// TIA Portal V20 export
Screen "190FX1Layout_Docking"  1276x673
  ScreenItem "Line_Header_X0_Y64" at 0,64 size 1276x0  Type=HmiLine
  ScreenItem "permanentareaborderrectangle" at 0,0 size 0x0  Type=HmiRectangle
  ScreenItem "Button_Back" at 2,2 size 90x60  Type=HmiButton
  ScreenItem "Move_Legend" at 1183,2 size 90x60  Type=HmiButton
  ScreenItem "Fusszeile_Button_ManualOPMode1_2" at 188,2 size 90x60  Type=HmiButton
  ScreenItem "文本域_22" at 1130,495 size 104x23  Type=HmiTextBox
  ScreenItem "面板容器_23" at 1177,528 size 96x32  Type=HmiFaceplateContainer
  ScreenItem "面板容器_22" at 1067,528 size 96x32  Type=HmiFaceplateContainer
  ScreenItem "面板容器_2" at 1091,4 size 88x58  Type=HmiFaceplateContainer
  ScreenItem "OPMode1_Blocked" at 1165,6 size 14x14  Type=HmiGraphicView
  ScreenItem "OPMode4_Foreground_Blocked" at 1091,4 size 88x58  Type=HmiGraphicView
  ScreenItem "Fusszeile_Button_ManualOPMode1_1" at 95,2 size 90x60  Type=HmiButton
  ScreenItem "LSicar_Valve8Pos_LeftHomeRightWork_WithPB_3" at 1099,110 size 160x53  Type=HmiFaceplateContainer
  ScreenItem "文本域_5" at 1107,83 size 139x22  Type=HmiTextBox
  ScreenItem "面板容器_15" at 54,347 size 65x43  Type=HmiFaceplateContainer
  ScreenItem "Graphic view_1" at 114,71 size 766x527  Type=HmiGraphicView
  ScreenItem "Line_4" at 527,411 size 146x156  Type=HmiLine
  ScreenItem "Line_5" at 509,439 size 5x185  Type=HmiLine
  ScreenItem "Line_6" at 104,365 size 253x0  Type=HmiLine
  ScreenItem "Line_7" at 406,338 size 1x280  Type=HmiLine
  ScreenItem "面板容器_13" at 613,609 size 142x51  Type=HmiFaceplateContainer
  ScreenItem "面板容器_12" at 312,609 size 142x51  Type=HmiFaceplateContainer
  ScreenItem "Faceplate container_5" at 483,609 size 65x43  Type=HmiFaceplateContainer
  ScreenItem "文本域_19" at 34,328 size 100x20  Type=HmiTextBox
  ScreenItem "文本域_6" at 312,567 size 140x40  Type=HmiTextBox
  ScreenItem "文本域_8" at 1172,-248 size 100x20  Type=HmiTextBox
  ScreenItem "文本域_9" at 1741,-563 size 100x20  Type=HmiTextBox
  ScreenItem "文本域_10" at 2310,-878 size 100x20  Type=HmiTextBox
  ScreenItem "文本域_11" at 462,587 size 100x20  Type=HmiTextBox
  ScreenItem "文本域_12" at 321,1215 size 100x20  Type=HmiTextBox
  ScreenItem "文本域_14" at 604,567 size 140x40  Type=HmiTextBox
  ScreenItem "Title_ScreenOverview_X390_Y2_1" at 384,2 size 510x57  Type=HmiTextBox
  ScreenItem "Button_Back_1" at 1180,606 size 90x60  Type=HmiButton
  ScreenItem "文本域_1" at -1,82 size 120x40  Type=HmiTextBox
  ScreenItem "文本域_27" at -1,126 size 120x40  Type=HmiTextBox
